(* IEC 61131-3 sources: kns-pump-station/tests/POUs/Station/FB_PumpProtection_Test, 11 files *)

(* ---- CurrentAtThresholdIsNotUnderload.method.decl.st ---- *)
// 04 §10.3: ток ровно 12 А — не недогрузка (строго меньше порога)
METHOD PRIVATE CurrentAtThresholdIsNotUnderload
VAR
    fbDut  : FB_PumpProtection;         // ФБ под тестом
    fbTime : PL.FB_FakeTime;            // подменное время, старт 1 ч
    stCfg  : ST_StationCfg;             // уставки по умолчанию: 12 А, 80 %, 15 с
END_VAR

(* ---- DisabledWhenThresholdZero.method.decl.st ---- *)
// 04 §18.2 № 28: rUnderload_A = 0 — контроль выключен
METHOD PRIVATE DisabledWhenThresholdZero
VAR
    fbDut  : FB_PumpProtection;         // ФБ под тестом
    fbTime : PL.FB_FakeTime;            // подменное время, старт 1 ч
    stCfg  : ST_StationCfg;             // уставки по умолчанию: 12 А, 80 %, 15 с
END_VAR

(* ---- NoUnderloadBelowMinSpeed.method.decl.st ---- *)
// 04 §10.3: частота ниже rUnderloadSpeed_pct — контроля нет; ровно 80 % — контроль есть (граница включительно)
METHOD PRIVATE NoUnderloadBelowMinSpeed
VAR
    fbDut  : FB_PumpProtection;         // ФБ под тестом
    fbTime : PL.FB_FakeTime;            // подменное время, старт 1 ч
    stCfg  : ST_StationCfg;             // уставки по умолчанию: 12 А, 80 %, 15 с
    fbDut2 : FB_PumpProtection;        // второй экземпляр: ровно 80 %
END_VAR

(* ---- NoUnderloadWhenCurrentInvalid.method.decl.st ---- *)
// 04 §10.3, PMI-29: ток недостоверен (нет связи) или не конечен — контроля недогрузки нет
METHOD PRIVATE NoUnderloadWhenCurrentInvalid
VAR
    fbDut  : FB_PumpProtection;         // ФБ под тестом
    fbTime : PL.FB_FakeTime;            // подменное время, старт 1 ч
    stCfg  : ST_StationCfg;             // уставки по умолчанию: 12 А, 80 %, 15 с
    uBits  : PL.U_RealBits;            // сборка NaN по битам
END_VAR

(* ---- OverheatInterlockWhileActive.method.decl.st ---- *)
// 04 §10.4, PMI-16: перегрев обмотки — бит KNS_ILK_OVERHEAT, пока сигнал активен, без фиксации
METHOD PRIVATE OverheatInterlockWhileActive
VAR
    fbDut  : FB_PumpProtection;         // ФБ под тестом
    fbTime : PL.FB_FakeTime;            // подменное время, старт 1 ч
    stCfg  : ST_StationCfg;             // уставки по умолчанию: 12 А, 80 %, 15 с
END_VAR

(* ---- ResetClearsLatch.method.decl.st ---- *)
// 04 §9.2: импульс сброса (фейсплейт, HS501, «Сбросить все») снимает фиксацию; отсчёт после сброса — заново
METHOD PRIVATE ResetClearsLatch
VAR
    fbDut  : FB_PumpProtection;         // ФБ под тестом
    fbTime : PL.FB_FakeTime;            // подменное время, старт 1 ч
    stCfg  : ST_StationCfg;             // уставки по умолчанию: 12 А, 80 %, 15 с
END_VAR

(* ---- Run.method.decl.st ---- *)
// Помощник: uiSteps шагов по 1 с; входы ФБ тест задаёт присваиванием
METHOD PRIVATE Run
VAR_IN_OUT
    fbDut  : FB_PumpProtection;         // ФБ под тестом
    fbTime : PL.FB_FakeTime;            // подменное время
    stCfg  : ST_StationCfg;             // уставки
END_VAR
VAR_INPUT
    uiSteps : UINT;                     // шагов по 1 с
END_VAR
VAR
    uiStep : UINT;                      // номер шага
END_VAR

(* ---- Run.method.impl.st ---- *)
FOR uiStep := 1 TO uiSteps DO
    fbTime.Advance(tStep := T#1S);
    fbDut(xReset := FALSE, itfTime := fbTime, stCfg := stCfg);
END_FOR

(* ---- TimeBackwardsRestartsUnderload.method.decl.st ---- *)
// Время назад — выдержка tUnderload начинается заново, ложной фиксации нет
METHOD PRIVATE TimeBackwardsRestartsUnderload
VAR
    fbDut  : FB_PumpProtection;         // ФБ под тестом
    fbTime : PL.FB_FakeTime;            // подменное время, старт 1 ч
    stCfg  : ST_StationCfg;             // уставки по умолчанию: 12 А, 80 %, 15 с
END_VAR

(* ---- UnderloadLatchedUntilReset.method.decl.st ---- *)
// 04 §10.3, PMI-15: фиксация держится, когда насос остановлен и ток вернулся, — до сброса насоса
METHOD PRIVATE UnderloadLatchedUntilReset
VAR
    fbDut  : FB_PumpProtection;         // ФБ под тестом
    fbTime : PL.FB_FakeTime;            // подменное время, старт 1 ч
    stCfg  : ST_StationCfg;             // уставки по умолчанию: 12 А, 80 %, 15 с
END_VAR

(* ---- UnderloadTripsAfterTUnderload.method.decl.st ---- *)
// 04 §10.3, PMI-15: ток ниже 12 А на частоте не ниже 80 % дольше tUnderload = 15 с — фиксация недогрузки и бит
// KNS_ILK_UNDERLOAD, не раньше
METHOD PRIVATE UnderloadTripsAfterTUnderload
VAR
    fbDut  : FB_PumpProtection;         // ФБ под тестом
    fbTime : PL.FB_FakeTime;            // подменное время, старт 1 ч
    stCfg  : ST_StationCfg;             // уставки по умолчанию: 12 А, 80 %, 15 с
END_VAR
